TYPE UDP_DATA : ARRAY[1..SIZEOF(S_TURBINECMD)*c_nNumTurbines] OF BYTE; END_TYPE

(* stored: Version 1.1.0.1
   DUT UDP_DATA: Id {0f72b5d4-758d-47da-9ab6-ac9e224924fa} *)
